Fanuc KAREL source: kt00331.KL

-- PROVISIONAL review KL for V770-1; original PC SHA256 2780378f876c86b62296e4fd973b0ab13b3633b59ae40756035f6d5c071377a3
-- Incomplete behavior may be omitted. Consult companion uncertainty JSON. Do not deploy.
PROGRAM KT00331
%NOLOCKGROUP
VAR
  I1 : INTEGER
  OUT : BOOLEAN
-- UNRESOLVED_DECL Y2 type=002018
BEGIN
  -- UNRESOLVED_PC offsets 5-16; opcodes 2E,23
  -- UNRESOLVED_PC offsets 21-35; opcodes 2E,22,9D,33,B2
  -- UNRESOLVED_PC offsets 40-62; opcodes 21,22,9D,33,B1,59,23
  -- UNRESOLVED_PC offsets 67-71; opcodes 7F
END KT00331
